// TIA Portal V18 export
DATA_BLOCK "DB_HMI_Data"   // DB1
{ S7_Optimized_Access := 'TRUE' }
// stored: MemoryReserve 100
   VAR
      motorForwardOn : Bool;
      motorReversOn : Bool;
      motorStop : Bool;
      frequencySetpoint : Real;
      frequencyActual : Real;
      voltageOut : Real;
      currentOut : Real;
      MinValueClamp : Int;
      MaxValueClamp : Int;
      frequencySource : Int;
      sensorOn : Bool;
      timerDelayMotorSensorsOn : Time;
      plcOnline : Bool;
      vfdOnline : Bool;
   END_VAR
BEGIN
END_DATA_BLOCK
